// TIA Portal V17 export
// export: Created 2000-01-01T00:00:00.0000000Z, ExportSetting None
TagTable "Water_HMI_IO"
  M1Pump : Bool  (PLC tag M1Pump, HMI_Connection_1, 100 ms)
  M1Valve : Bool  (PLC tag M1Valve, HMI_Connection_1, 100 ms)
  M1Reset : Bool  (PLC tag M1Reset, HMI_Connection_1, 100 ms)
  M1PumpFlow : Bool  (PLC tag M1PumpFlow, HMI_Connection_1, 100 ms)
  M1ValveFlow : Bool  (PLC tag M1ValveFlow, HMI_Connection_1, 100 ms)
  M1MixerRun : Bool  (PLC tag M1MixerRun, HMI_Connection_1, 100 ms)
  M2Pump : Bool  (PLC tag M2Pump, HMI_Connection_1, 100 ms)
  M2V1 : Bool  (PLC tag M2V1, HMI_Connection_1, 100 ms)
  M2V2 : Bool  (PLC tag M2V2, HMI_Connection_1, 100 ms)
  M2V3 : Bool  (PLC tag M2V3, HMI_Connection_1, 100 ms)
  M2Reset : Bool  (PLC tag M2Reset, HMI_Connection_1, 100 ms)
  M2PumpFlow : Bool  (PLC tag M2PumpFlow, HMI_Connection_1, 100 ms)
  M2Irrigate : Bool  (PLC tag M2Irrigate, HMI_Connection_1, 100 ms)
  M2Reaction : Bool  (PLC tag M2Reaction, HMI_Connection_1, 100 ms)
  M2LoadFlow : Bool  (PLC tag M2LoadFlow, HMI_Connection_1, 100 ms)
  M2TruckMoving : Bool  (PLC tag M2TruckMoving, HMI_Connection_1, 100 ms)
  M1Tank : Int  (PLC tag M1Tank, HMI_Connection_1, 100 ms)
  M1Pond : Int  (PLC tag M1Pond, HMI_Connection_1, 100 ms)
  M1MixFrame : Int  (PLC tag M1MixFrame, HMI_Connection_1, 100 ms)
  M2Reservoir : Int  (PLC tag M2Reservoir, HMI_Connection_1, 100 ms)
  M2Tank : Int  (PLC tag M2Tank, HMI_Connection_1, 100 ms)
  M2Truck : Int  (PLC tag M2Truck, HMI_Connection_1, 100 ms)
  M2TruckPosition : Int  (PLC tag M2TruckPosition, HMI_Connection_1, 100 ms)
  M2GrassTotal : Int  (PLC tag M2GrassTotal, HMI_Connection_1, 100 ms)
  M1PumpFrame : Int  (PLC tag M1PumpFrame, HMI_Connection_1, 100 ms)
  M1ValveFrame : Int  (PLC tag M1ValveFrame, HMI_Connection_1, 100 ms)
  M2PumpFrame : Int  (PLC tag M2PumpFrame, HMI_Connection_1, 100 ms)
  M2V1Frame : Int  (PLC tag M2V1Frame, HMI_Connection_1, 100 ms)
  M2V2Frame : Int  (PLC tag M2V2Frame, HMI_Connection_1, 100 ms)
  M2V3Frame : Int  (PLC tag M2V3Frame, HMI_Connection_1, 100 ms)
